Fanuc KAREL source: KD00023.KL

PROGRAM KD00023
%NOLOCKGROUP
VAR
  I: INTEGER
  J: INTEGER
  B: BOOLEAN
  R: REAL
  S: STRING[80]
  SAVED IN DRAM: INTEGER
BEGIN
  I = SAVED
END KD00023
